RESOURCE RES0 : EMB_RES_ECO
  FBS
    MGE_LODO : MGE_Generico(cfgTempoCom := 5);
    MGE_DESINFECCAO : MGE_Generico(cfgTempoCom := 5);
    DESINFECCAO : Desinfeccao_UV;
    DESINF_A2_DI32K0 : IO_DI32(WORD0 := '$${PATH}DESINF_A2_DI32K_WORD0', WORD1 := '$${PATH}DESINF_A2_DI32K_WORD1', CONN := '$${PATH}DESINF_A2_DI32K0_CONN', COM_OK := 'RES0.DESINFECCAO.stsRemotaComOk', DI_0 := 'RES0.DESINFECCAO.djPCEDesligado', DI_1 := 'RES0.DESINFECCAO.djPCMDesligado', DI_2 := 'RES0.DESINFECCAO.djUV01', DI_3 := 'RES0.DESINFECCAO.djUV02', DI_4 := 'RES0.DESINFECCAO.djVC01', DI_5 := 'RES0.DESINFECCAO.djMO01');
    DesidratacaoLodo : DesidratacaoLodo;
    EstocagemLodo : EstocagemLodo;
    LODO_A3_DI32K0 : IO_DI32(WORD0 := '$${PATH}LODO_A3_DI32K_WORD0', WORD1 := '$${PATH}LODO_A3_DI32K_WORD1', CONN := '$${PATH}LODO_R1_CONN', COM_OK := 'RES0.DesidratacaoLodo.stsRemota1ComOk', DI_0 := 'RES0.DesidratacaoLodo.djPCE', DI_1 := 'RES0.DesidratacaoLodo.stsEmergenciaPainel', DI_2 := 'RES0.DesidratacaoLodo.djPCM', DI_3 := 'RES0.DesidratacaoLodo.djSO01', DI_4 := 'RES0.EstocagemLodo.SO_900_01.stsLocal', DI_5 := 'RES0.EstocagemLodo.SO_900_01.stsRemoto', DI_6 := 'RES0.EstocagemLodo.SO_900_01.stsLigado', DI_7 := 'RES0.EstocagemLodo.SO_900_01.stsSemFalha', DI_8 := 'RES0.DesidratacaoLodo.djSO02', DI_9 := 'RES0.EstocagemLodo.SO_900_02.stsLocal', DI_10 := 'RES0.EstocagemLodo.SO_900_02.stsRemoto', DI_11 := 'RES0.EstocagemLodo.SO_900_02.stsLigado', DI_12 := 'RES0.EstocagemLodo.SO_900_02.stsSemFalha', DI_13 := 'RES0.DesidratacaoLodo.djAD01', DI_14 := 'RES0.DesidratacaoLodo.djAD02', DI_15 := 'RES0.DesidratacaoLodo.djAD03', DI_16 := 'RES0.DesidratacaoLodo.djPP01', DI_17 := 'RES0.DesidratacaoLodo.djMN01', DI_18 := 'RES0.DesidratacaoLodo.djMN02', DI_19 := 'RES0.DesidratacaoLodo.djMN03', DI_20 := 'RES0.DesidratacaoLodo.djMN04', DI_21 := 'RES0.DesidratacaoLodo.djMN05', DI_22 := 'RES0.DesidratacaoLodo.djBO01', DI_23 := 'RES0.DesidratacaoLodo.BO_900_01.stsLocal', DI_24 := 'RES0.DesidratacaoLodo.BO_900_01.stsRemoto', DI_25 := 'RES0.DesidratacaoLodo.BO_900_01.stsLigado', DI_26 := 'RES0.DesidratacaoLodo.BO_900_01.stsSemFalha', DI_27 := 'RES0.DesidratacaoLodo.BO_900_01.stsProtecaoTermica', DI_28 := 'RES0.DesidratacaoLodo.djBO02', DI_29 := 'RES0.DesidratacaoLodo.BO_900_02.stsLocal', DI_30 := 'RES0.DesidratacaoLodo.BO_900_02.stsRemoto', DI_31 := 'RES0.DesidratacaoLodo.BO_900_02.stsLigado');
    LODO_A4_DI32K0 : IO_DI32(WORD0 := '$${PATH}LODO_A4_DI32K_WORD0', WORD1 := '$${PATH}LODO_A4_DI32K_WORD1', CONN := 'RES0.LODO_A3_DI32K0.LODO_R1_CONN', DI_0 := 'RES0.DesidratacaoLodo.BO_900_02.stsSemFalha', DI_1 := 'RES0.DesidratacaoLodo.BO_900_02.stsProtecaoTermica', DI_2 := 'RES0.DesidratacaoLodo.djBO03', DI_3 := 'RES0.DesidratacaoLodo.BO_900_03.stsLocal', DI_4 := 'RES0.DesidratacaoLodo.BO_900_03.stsRemoto', DI_5 := 'RES0.DesidratacaoLodo.BO_900_03.stsLigado', DI_6 := 'RES0.DesidratacaoLodo.BO_900_03.stsSemFalha', DI_7 := 'RES0.DesidratacaoLodo.BO_900_03.stsProtecaoTermica', DI_8 := 'RES0.DesidratacaoLodo.djBR01', DI_9 := 'RES0.DesidratacaoLodo.BR_900_01.stsLocal', DI_10 := 'RES0.DesidratacaoLodo.BR_900_01.stsRemoto', DI_11 := 'RES0.DesidratacaoLodo.BR_900_01.stsLigado', DI_12 := 'RES0.DesidratacaoLodo.BR_900_01.stsSemFalha', DI_13 := 'RES0.DesidratacaoLodo.stsMonitTrafo', DI_14 := 'RES0.DesidratacaoLodo.djBR02', DI_15 := 'RES0.DesidratacaoLodo.BR_900_02.stsLocal', DI_16 := 'RES0.DesidratacaoLodo.BR_900_02.stsRemoto', DI_17 := 'RES0.DesidratacaoLodo.BR_900_02.stsLigado', DI_18 := 'RES0.DesidratacaoLodo.BR_900_02.stsSemFalha', DI_19 := 'RES0.DesidratacaoLodo.stsMonitFonte', DI_20 := 'RES0.DesidratacaoLodo.djVA01', DI_21 := 'RES0.DesidratacaoLodo.djVA02', DI_22 := 'RES0.DesidratacaoLodo.djVE01', DI_23 := 'RES0.DesidratacaoLodo.djVE02', DI_25 := 'RES0.DesidratacaoLodo.djVA06', DI_26 := 'RES0.DesidratacaoLodo.djVA07', DI_27 := 'RES0.DesidratacaoLodo.djVA08', DI_28 := 'RES0.DesidratacaoLodo.djVA09', DI_29 := 'RES0.DesidratacaoLodo.djVA10', DI_30 := 'RES0.DesidratacaoLodo.djVA11', DI_31 := 'RES0.DesidratacaoLodo.djVA12');
    LODO_A5_DI32K0 : IO_DI32(WORD0 := '$${PATH}LODO_A5_DI32K_WORD0', WORD1 := '$${PATH}LODO_A5_DI32K_WORD1', CONN := 'RES0.LODO_A3_DI32K0.LODO_R1_CONN', DI_0 := 'RES0.DesidratacaoLodo.djVA13', DI_1 := 'RES0.DesidratacaoLodo.djVB03', DI_2 := 'RES0.DesidratacaoLodo.djVB04');
    LODO_A7_DQ32TK0 : IO_DQ32(WORD0 := '$${PATH}LODO_A7_DQ32TK_WORD0', WORD1 := '$${PATH}LODO_A7_DQ32TK_WORD1', CONN := 'RES0.LODO_A3_DI32K0.LODO_R1_CONN', DO_0 := 'RES0.EstocagemLodo.SO_900_01.cmdAcionamento', DO_1 := 'RES0.EstocagemLodo.SO_900_01.cmdReset', DO_2 := 'RES0.EstocagemLodo.SO_900_02.cmdAcionamento', DO_3 := 'RES0.EstocagemLodo.SO_900_02.cmdReset', DO_4 := 'RES0.DesidratacaoLodo.BO_900_01.cmdAcionamento', DO_5 := 'RES0.DesidratacaoLodo.BO_900_01.cmdReset', DO_6 := 'RES0.DesidratacaoLodo.BO_900_02.cmdAcionamento', DO_7 := 'RES0.DesidratacaoLodo.BO_900_02.cmdReset', DO_8 := 'RES0.DesidratacaoLodo.BO_900_03.cmdAcionamento', DO_9 := 'RES0.DesidratacaoLodo.BO_900_03.cmdReset', DO_10 := 'RES0.DesidratacaoLodo.BR_900_01.cmdAcionamento', DO_11 := 'RES0.DesidratacaoLodo.BR_900_01.cmdReset', DO_12 := 'RES0.DesidratacaoLodo.BR_900_02.cmdAcionamento', DO_13 := 'RES0.DesidratacaoLodo.BR_900_02.cmdReset', DO_14 := 'RES0.DesidratacaoLodo.cmdSV01', DO_15 := 'RES0.DesidratacaoLodo.cmdSV02', DO_16 := 'RES0.DesidratacaoLodo.cmdSV03', DO_17 := 'RES0.DesidratacaoLodo.cmdSV04', DO_18 := 'RES0.DesidratacaoLodo.cmdSV06', DO_19 := 'RES0.DesidratacaoLodo.cmdSV08');
    SR_LODO_A2_REMOTA1 : Status_Remota;
    SR_LODO_A10_REMOTA2 : Status_Remota;
    SR_DESINF_A1_REMOTA : Status_Remota;
    DPAC_FULLINIT1 : DPAC_FULLINIT;
  END_FBS
  EVENT_CONNECTIONS
    START.COLD TO DPAC_FULLINIT1.INIT;
    START.WARM TO DPAC_FULLINIT1.INIT;
    START.ONLINECHANGE TO DPAC_FULLINIT1.OC_RETRIGGER;
    EstocagemLodo.974B4969DB603762 TO DesidratacaoLodo.91E17855232378A8;
    EstocagemLodo.E3809710B35A5BE3 TO DesidratacaoLodo.335836E160C77742;
    DesidratacaoLodo.D64A39BCF02DDEB2 TO EstocagemLodo.AB5FAE61D1BCDDFE;
    DesidratacaoLodo.EA9A2427D178E8B5 TO EstocagemLodo.39F3DF7DDD7B4C23;
    DesidratacaoLodo.EE8958653A86D261 TO EstocagemLodo.4FA8CBCB1032FBD8;
  END_CONNECTIONS
  DATA_CONNECTIONS
    DesidratacaoLodo.9DCD88E1901DA328 TO EstocagemLodo.A8767255ECC4E3FD;
    EstocagemLodo.649314760363E488 TO DesidratacaoLodo.AC99B8EE5C6DBA64;
    EstocagemLodo.B87FCF9EF6E17A10 TO DesidratacaoLodo.D231A14376C3E2F6;
    EstocagemLodo.273D781A989DEA3F TO DesidratacaoLodo.DE00033B699DACF0;
    EstocagemLodo.0D2CE8145A8A40C5 TO DesidratacaoLodo.099E44A540EF9490;
    EstocagemLodo.E7A1F2C70FD2876B TO DesidratacaoLodo.426B37B9A495B79C;
    EstocagemLodo.5C0EE27FAC026E42 TO DesidratacaoLodo.FD17B98D889E4E9C;
    EstocagemLodo.28C5117F80A71252 TO DesidratacaoLodo.91FA512D1B0CCA17;
    EstocagemLodo.F39C9B782425030B TO DesidratacaoLodo.18A2A222BB911413;
    EstocagemLodo.CA5C991A51FB83CF TO DesidratacaoLodo.14561E73765FBECA;
    EstocagemLodo.5405EB7088EC4BDE TO DesidratacaoLodo.1CD77F0C67EACF01;
    DesidratacaoLodo.317BB96205F3F911 TO EstocagemLodo.EE49B187C469C0B7;
    DesidratacaoLodo.A2D8149F0FE69321 TO EstocagemLodo.E59CBDC75C3131D4;
    DesidratacaoLodo.08464482A0BF6120 TO EstocagemLodo.8E87331950BD000E;
    DesidratacaoLodo.4080C84A5DF2BAE8 TO EstocagemLodo.3B31F82669E06299;
  END_CONNECTIONS
END_RESOURCE
